DATA_BLOCK "PressDemo"
{ S7_Optimized_Access := 'TRUE' }
VERSION : 0.1
NON_RETAIN
"FB_PressDemoUnit"
BEGIN
END_DATA_BLOCK
